GLOBALCONSTANTS TestConstants (* Global constants for import export tests *)
  (* Standard: 61499-1; Description: Copyright (c) 2026 Martin Erich Jobst This program and the accompanying materials are made available under the terms of the Eclipse Public License 2.0 which is available at https://www.eclipse.org/legal/epl-2.0/ SPDX-License-Identifier: EPL-2.0 *)
  (* Version 1.0, 2026-10-23, Martin Jobst *)
  {SET_ATTRIBUTE(IntegerAttribute, 10)}
  VAR_GLOBAL CONSTANT
    ANSWER : DINT := DINT#42; (* Answer *)
  END_VAR
END_GLOBALCONSTANTS
